(* IEC 61131-3 sources: llm-plc-st-eval/data/calibracion/gpt-4o-2024-08-06/B1/few_shot, 3 files *)

(* ---- ejec_1.st ---- *)
```pascal
FUNCTION_BLOCK FB_Motor
VAR_INPUT
    btnMarcha : BOOL; (* Botón de marcha *)
    btnParo : BOOL;   (* Botón de paro *)
    btnEmerg : BOOL;  (* Botón de paro de emergencia *)
END_VAR
VAR_OUTPUT
    motorOn : BOOL;   (* Estado del motor *)
END_VAR
VAR
    motorLatch : BOOL; (* Latch para mantener el motor encendido *)
END_VAR

(* Control de arranque y paro del motor *)
IF btnEmerg THEN
    motorLatch := FALSE; (* Paro de emergencia, el motor no puede rearrancar *)
ELSIF btnParo THEN
    motorLatch := FALSE; (* Paro normal, apaga el motor *)
ELSIF btnMarcha THEN
    motorLatch := TRUE;  (* Arranca el motor y lo mantiene encendido *)
END_IF

motorOn := motorLatch; (* Actualiza el estado del motor *)
END_FUNCTION_BLOCK
```

(* ---- ejec_2.st ---- *)
```pascal
FUNCTION_BLOCK FB_Motor
VAR_INPUT
    btnMarcha : BOOL; (* Botón de marcha *)
    btnParo : BOOL;   (* Botón de paro *)
    btnEmerg : BOOL;  (* Botón de paro de emergencia *)
END_VAR
VAR_OUTPUT
    motorOn : BOOL;   (* Estado del motor *)
END_VAR
VAR
    motorActivo : BOOL; (* Estado interno del motor *)
END_VAR

(* Lógica de control del motor *)
IF btnEmerg THEN
    motorActivo := FALSE; (* Paro de emergencia, desactiva el motor *)
ELSIF btnParo THEN
    motorActivo := FALSE; (* Botón de paro, desactiva el motor *)
ELSIF btnMarcha THEN
    motorActivo := TRUE;  (* Botón de marcha, activa el motor *)
END_IF

motorOn := motorActivo; (* Salida del estado del motor *)
END_FUNCTION_BLOCK
```

(* ---- ejec_3.st ---- *)
```pascal
FUNCTION_BLOCK FB_Motor
VAR_INPUT
    btnMarcha : BOOL; (* Botón de marcha *)
    btnParo : BOOL;   (* Botón de paro *)
    btnEmerg : BOOL;  (* Botón de paro de emergencia *)
END_VAR
VAR_OUTPUT
    motorOn : BOOL;   (* Estado del motor *)
END_VAR
VAR
    motorActivo : BOOL; (* Estado interno del motor *)
END_VAR

(* Lógica de control del motor *)
IF btnEmerg THEN
    motorActivo := FALSE; (* Paro de emergencia desactiva el motor *)
ELSIF btnParo THEN
    motorActivo := FALSE; (* Botón de paro desactiva el motor *)
ELSIF btnMarcha THEN
    motorActivo := TRUE;  (* Botón de marcha activa el motor *)
END_IF

motorOn := motorActivo; (* Salida del estado del motor *)
END_FUNCTION_BLOCK
```
